// TIA Portal V20 export
VAR_GLOBAL   // PLC tag table "PLC-A4-DQ"
   "-KA12" AT %Q8.0 : Bool;
   "-KA13" AT %Q8.1 : Bool;
   "-KA14" AT %Q8.2 : Bool;
   "-KA15" AT %Q8.3 : Bool;
   "-KA16" AT %Q8.4 : Bool;
   "-KA17" AT %Q8.5 : Bool;
   RESERVE_DQ_ AT %Q8.6 : Bool;
   RESERVE_DQ_1 AT %Q8.7 : Bool;
   RESERVE_DQ_2 AT %Q9.0 : Bool;   // vyrazovac
   RESERVE_DQ_3 AT %Q9.1 : Bool;
   RESERVE_DQ_4 AT %Q9.2 : Bool;
   RESERVE_DQ_5 AT %Q9.3 : Bool;
   RESERVE_DQ_6 AT %Q9.4 : Bool;
   RESERVE_DQ_7 AT %Q9.5 : Bool;
   RESERVE_DQ_8 AT %Q9.6 : Bool;
   RESERVE_DQ_9 AT %Q9.7 : Bool;
END_VAR
